(* IEC 61131-3 sources: OpenPLC_v3_afl_compile/webserver/st_files, 3 files *)

(* ---- blank_program.st ---- *)
PROGRAM prog0
  VAR
    var_in : BOOL;
    var_out : BOOL;
  END_VAR

  var_out := var_in;
END_PROGRAM

CONFIGURATION Config0

  RESOURCE Res0 ON PLC
    TASK Main(INTERVAL := T#50ms,PRIORITY := 0);
    PROGRAM Inst0 WITH Main : prog0;
  END_RESOURCE
END_CONFIGURATION

(* ---- water_tank_simple.st ---- *)
PROGRAM water_tank
  VAR
    tank_level AT %QW0 : INT := 500;
    pump_state AT %QW1 : INT := 0;
    alarm_state AT %QW2 : INT := 0;
    setpoint AT %QW3 : INT := 500;
  END_VAR

  IF pump_state = 1 THEN
    tank_level := tank_level + 5;
  END_IF;

  IF tank_level > 0 THEN
    tank_level := tank_level - 2;
  END_IF;

  IF tank_level > 1000 THEN
    tank_level := 1000;
  END_IF;

  IF tank_level < 0 THEN
    tank_level := 0;
  END_IF;

  IF tank_level < 300 THEN
    pump_state := 1;
  END_IF;

  IF tank_level > 700 THEN
    pump_state := 0;
  END_IF;

  IF tank_level > 850 THEN
    alarm_state := 1;
  END_IF;

  IF tank_level < 800 THEN
    alarm_state := 0;
  END_IF;

END_PROGRAM

CONFIGURATION Config0
  RESOURCE Res0 ON PLC
    TASK task0(INTERVAL := T#20ms,PRIORITY := 0);
    PROGRAM instance0 WITH task0 : water_tank;
  END_RESOURCE
END_CONFIGURATION

(* ---- webserver_program.st ---- *)
PROGRAM prog0
  VAR
    var_in : BOOL;
    var_out : BOOL;
  END_VAR

  var_out := var_in;
END_PROGRAM

CONFIGURATION Config0

  RESOURCE Res0 ON PLC
    TASK Main(INTERVAL := T#50ms,PRIORITY := 0);
    PROGRAM Inst0 WITH Main : prog0;
  END_RESOURCE
END_CONFIGURATION
